// TwinCAT 3 PLC project TestFrameworkPLC
// ProgramVersion: 3.1.4026.28
// libraries:
//   [IO_ReadWrite], * (BACA_Apps)
//   Tc2_Standard, * (Beckhoff Automation GmbH)
//   Tc2_System, * (Beckhoff Automation GmbH)
//   Tc3_PlcTestFramework, * (Beckhoff Automation GmbH)
// project tree:
//   / PlcTask.TcTTO
//   POUs/ FB_IO_Test.TcPOU, MAIN.TcPOU
// (motion and I/O tree: see PLC project io_readwrite)
// real-time tasks:
//   TASK PlcTask1: cycle T#1ms, priority 21, ADS port 351
// variable links:
//   TestFrameworkPLC/TestFrameworkPLC Instance <-> Device 1 (EtherCAT)/Term 1 (EK1200)/Term 2 (EL1002)
//     PlcTask Inputs/MAIN.fbT1.fbIOtester.bIn <-> Channel 1/Input
//   TestFrameworkPLC/TestFrameworkPLC Instance <-> Device 1 (EtherCAT)/Term 1 (EK1200)/Term 3 (EL2002)
//     PlcTask Outputs/MAIN.fbT1.fbIOtester.bOut <-> Channel 1/Output

CONFIGURATION TestFrameworkPLC
    RESOURCE PLC ON TwinCAT3
        TASK PlcTask(INTERVAL := T#1ms, PRIORITY := 21);
        PROGRAM MAIN WITH PlcTask : MAIN;
    END_RESOURCE
END_CONFIGURATION

// ---- POUs/MAIN.TcPOU
PROGRAM MAIN
VAR
	fbT1 : FB_IO_Test;
END_VAR

Tc3_PlcTestFramework.F_CallTestController();

END_PROGRAM

// ---- POUs/FB_IO_Test.TcPOU
{ attribute 'Name':='...' }
{ attribute 'Timeout':='t#20s' }
{ attribute 'Owner':='BACA_Apps' }
{ attribute 'Category':='IO Check' }
FUNCTION_BLOCK FB_IO_Test EXTENDS FB_TestCaseBase
VAR_INPUT
END_VAR
VAR_OUTPUT
END_VAR
VAR
	fbIOtester : IO_ReadWrite.FB_IO_ReadWrite;			
END_VAR

fbIOtester.bExecute := TRUE; 
fbIOtester.timerDelay := T#100MS;

IF fbIOtester.bDone THEN
	AssertTrue(bCondition := fbIOtester.bHighMatch, sMessage := 'Channel 1 failed HIGH check');
	AssertTrue(bCondition := fbIOtester.bLowMatch, sMessage := 'Channel 1 failed LOW check');
	fbIOtester.bExecute := FALSE;
	Succeed();
END_IF

fbIOtester();

END_FUNCTION_BLOCK
